// TIA Portal V21 export
// export: Created 2026-11-10T19:21:33.6052919Z, ExportSetting WithDefaults, DisplayName Totally Integrated Automation Portal, DisplayVersion V21 Update 3, DisplayName STEP 7 Professional, DisplayVersion V21 Update 3, DisplayName STEP 7 Safety, DisplayVersion V21, DisplayName Tech WebApplication, DisplayVersion V21, DisplayName WinCC Basic/Comfort/Advanced, DisplayVersion V21 Update 3, DisplayName WinCC Unified, DisplayVersion V21 Update 3
FUNCTION_BLOCK "FB_Lad_us003"   // FB6, LAD
{ S7_Optimized_Access := 'TRUE' }
VERSION : 0.1
// stored: AutoNumber true, IsIECCheckEnabled false, IsRetainMemResEnabled false, MemoryReserve 100, SetENOAutomatically false, UDAEnableTagReadback false
   VAR_INPUT
      v_port : PORT;
      v_baud : DInt;
   END_VAR
   VAR_OUTPUT
      v_error : Bool;
      v_status : Word;
   END_VAR
   VAR_IN_OUT
      v_uss_db : P2P_USS_BASE;
   END_VAR
   VAR
      inst { S7_SetPoint := 'True'} : USS_Port_Scan;
   END_VAR
BEGIN

REGION Network 1: USS_PORT - Edit communication via USS network
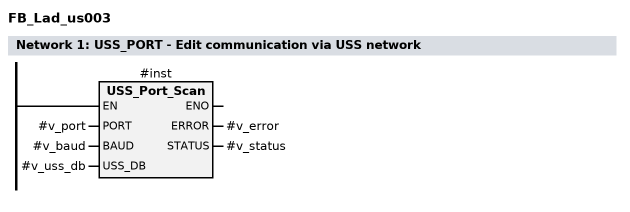
   RUNG wire#powerrail
      #inst.USS_Port_Scan(PORT := #v_port, BAUD := #v_baud, USS_DB := #v_uss_db, ERROR => #v_error, STATUS => #v_status)
   END_RUNG
   // the same network as SCL:
   #inst(PORT := #v_port, BAUD := #v_baud, USS_DB := #v_uss_db, ERROR => #v_error, STATUS => #v_status);   // USS_Port_Scan
END_REGION
END_FUNCTION_BLOCK
